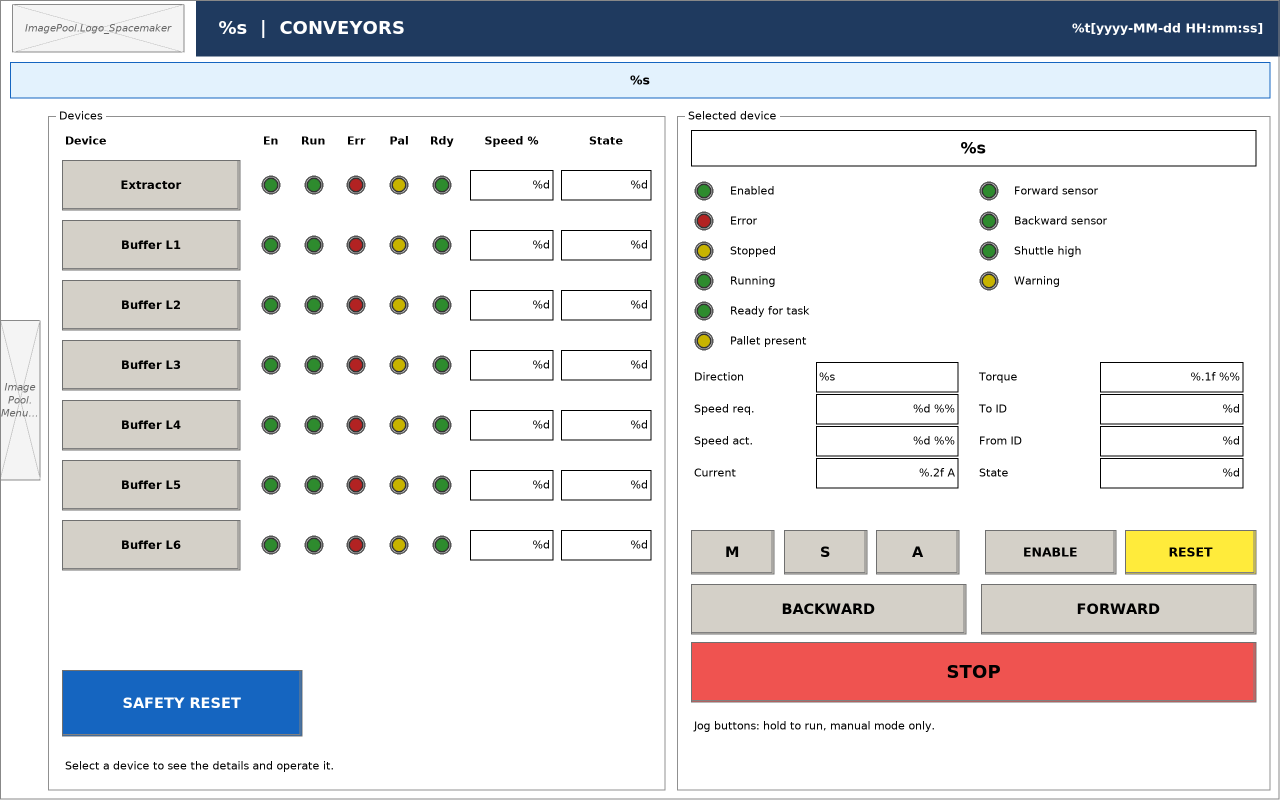
VISUALIZATION CNV  // 1280x800
    Rectangle (0,0 196x56)
        OnMouseClick: change screen: Main
    Image (12,4 172x48), image: ImagePool.Logo_Spacemaker
        OnMouseClick: change screen: Main
    Rectangle (196,0 1084x56), "%s | CONVEYORS", text variable: GVL_HMI_System.stStatus.sSystemName
    Rectangle (930,8 336x40), "%t[yyyy-MM-dd HH:mm:ss]", text variable: GVL_HMI_System.stStatus.dtNow
    Rectangle (10,62 1260x36), "%s", text variable: GVL_HMI_System.stStatus.sMessage, colour toggle: GVL_HMI_System.stStatus.bMessageAlarm
    GroupBox (48,108 617x682), "Devices"
    Rectangle (62,128 178x26), "Device"
    Rectangle (250,128 42x26), "En"
    Rectangle (292,128 43x26), "Run"
    Rectangle (335,128 43x26), "Err"
    Rectangle (378,128 43x26), "Pal"
    Rectangle (421,128 42x26), "Rdy"
    Rectangle (470,128 83x26), "Speed %"
    Rectangle (561,128 90x26), "State"
    Button (62,160 178x50), "Extractor", colour toggle: GVL_HMI_CNV.astConveyor[0].bSelected
        OnMouseClick: execute { GVL_HMI_CNV.uiSelected := 0; }
    Lamp1 (260,174 22x22), variable: GVL_HMI_CNV.astConveyor[0].bEnabled, style: Lamp-Lamp1-Green
    Lamp1 (303,174 22x22), variable: GVL_HMI_CNV.astConveyor[0].bRunning, style: Lamp-Lamp1-Green
    Lamp1 (345,174 22x22), variable: GVL_HMI_CNV.astConveyor[0].bError, style: Lamp-Lamp1-Red
    Lamp1 (388,174 22x22), variable: GVL_HMI_CNV.astConveyor[0].bOccupied, style: Lamp-Lamp1-Yellow
    Lamp1 (431,174 22x22), variable: GVL_HMI_CNV.astConveyor[0].bReadyForTask, style: Lamp-Lamp1-Green
    Rectangle (470,170 83x30), "%d", text variable: GVL_HMI_CNV.astConveyor[0].iSpeedActual_pct
    Rectangle (561,170 90x30), "%d", text variable: GVL_HMI_CNV.astConveyor[0].uiStateMachine
    Button (62,220 178x50), "Buffer L1", colour toggle: GVL_HMI_CNV.astConveyor[1].bSelected
        OnMouseClick: execute { GVL_HMI_CNV.uiSelected := 1; }
    Lamp1 (260,234 22x22), variable: GVL_HMI_CNV.astConveyor[1].bEnabled, style: Lamp-Lamp1-Green
    Lamp1 (303,234 22x22), variable: GVL_HMI_CNV.astConveyor[1].bRunning, style: Lamp-Lamp1-Green
    Lamp1 (345,234 22x22), variable: GVL_HMI_CNV.astConveyor[1].bError, style: Lamp-Lamp1-Red
    Lamp1 (388,234 22x22), variable: GVL_HMI_CNV.astConveyor[1].bOccupied, style: Lamp-Lamp1-Yellow
    Lamp1 (431,234 22x22), variable: GVL_HMI_CNV.astConveyor[1].bReadyForTask, style: Lamp-Lamp1-Green
    Rectangle (470,230 83x30), "%d", text variable: GVL_HMI_CNV.astConveyor[1].iSpeedActual_pct
    Rectangle (561,230 90x30), "%d", text variable: GVL_HMI_CNV.astConveyor[1].uiStateMachine
    Button (62,280 178x50), "Buffer L2", colour toggle: GVL_HMI_CNV.astConveyor[2].bSelected
        OnMouseClick: execute { GVL_HMI_CNV.uiSelected := 2; }
    Lamp1 (260,294 22x22), variable: GVL_HMI_CNV.astConveyor[2].bEnabled, style: Lamp-Lamp1-Green
    Lamp1 (303,294 22x22), variable: GVL_HMI_CNV.astConveyor[2].bRunning, style: Lamp-Lamp1-Green
    Lamp1 (345,294 22x22), variable: GVL_HMI_CNV.astConveyor[2].bError, style: Lamp-Lamp1-Red
    Lamp1 (388,294 22x22), variable: GVL_HMI_CNV.astConveyor[2].bOccupied, style: Lamp-Lamp1-Yellow
    Lamp1 (431,294 22x22), variable: GVL_HMI_CNV.astConveyor[2].bReadyForTask, style: Lamp-Lamp1-Green
    Rectangle (470,290 83x30), "%d", text variable: GVL_HMI_CNV.astConveyor[2].iSpeedActual_pct
    Rectangle (561,290 90x30), "%d", text variable: GVL_HMI_CNV.astConveyor[2].uiStateMachine
    Button (62,340 178x50), "Buffer L3", colour toggle: GVL_HMI_CNV.astConveyor[3].bSelected
        OnMouseClick: execute { GVL_HMI_CNV.uiSelected := 3; }
    Lamp1 (260,354 22x22), variable: GVL_HMI_CNV.astConveyor[3].bEnabled, style: Lamp-Lamp1-Green
    Lamp1 (303,354 22x22), variable: GVL_HMI_CNV.astConveyor[3].bRunning, style: Lamp-Lamp1-Green
    Lamp1 (345,354 22x22), variable: GVL_HMI_CNV.astConveyor[3].bError, style: Lamp-Lamp1-Red
    Lamp1 (388,354 22x22), variable: GVL_HMI_CNV.astConveyor[3].bOccupied, style: Lamp-Lamp1-Yellow
    Lamp1 (431,354 22x22), variable: GVL_HMI_CNV.astConveyor[3].bReadyForTask, style: Lamp-Lamp1-Green
    Rectangle (470,350 83x30), "%d", text variable: GVL_HMI_CNV.astConveyor[3].iSpeedActual_pct
    Rectangle (561,350 90x30), "%d", text variable: GVL_HMI_CNV.astConveyor[3].uiStateMachine
    Button (62,400 178x50), "Buffer L4", colour toggle: GVL_HMI_CNV.astConveyor[4].bSelected
        OnMouseClick: execute { GVL_HMI_CNV.uiSelected := 4; }
    Lamp1 (260,414 22x22), variable: GVL_HMI_CNV.astConveyor[4].bEnabled, style: Lamp-Lamp1-Green
    Lamp1 (303,414 22x22), variable: GVL_HMI_CNV.astConveyor[4].bRunning, style: Lamp-Lamp1-Green
    Lamp1 (345,414 22x22), variable: GVL_HMI_CNV.astConveyor[4].bError, style: Lamp-Lamp1-Red
    Lamp1 (388,414 22x22), variable: GVL_HMI_CNV.astConveyor[4].bOccupied, style: Lamp-Lamp1-Yellow
    Lamp1 (431,414 22x22), variable: GVL_HMI_CNV.astConveyor[4].bReadyForTask, style: Lamp-Lamp1-Green
    Rectangle (470,410 83x30), "%d", text variable: GVL_HMI_CNV.astConveyor[4].iSpeedActual_pct
    Rectangle (561,410 90x30), "%d", text variable: GVL_HMI_CNV.astConveyor[4].uiStateMachine
    Button (62,460 178x50), "Buffer L5", colour toggle: GVL_HMI_CNV.astConveyor[5].bSelected
        OnMouseClick: execute { GVL_HMI_CNV.uiSelected := 5; }
    Lamp1 (260,474 22x22), variable: GVL_HMI_CNV.astConveyor[5].bEnabled, style: Lamp-Lamp1-Green
    Lamp1 (303,474 22x22), variable: GVL_HMI_CNV.astConveyor[5].bRunning, style: Lamp-Lamp1-Green
    Lamp1 (345,474 22x22), variable: GVL_HMI_CNV.astConveyor[5].bError, style: Lamp-Lamp1-Red
    Lamp1 (388,474 22x22), variable: GVL_HMI_CNV.astConveyor[5].bOccupied, style: Lamp-Lamp1-Yellow
    Lamp1 (431,474 22x22), variable: GVL_HMI_CNV.astConveyor[5].bReadyForTask, style: Lamp-Lamp1-Green
    Rectangle (470,470 83x30), "%d", text variable: GVL_HMI_CNV.astConveyor[5].iSpeedActual_pct
    Rectangle (561,470 90x30), "%d", text variable: GVL_HMI_CNV.astConveyor[5].uiStateMachine
    Button (62,520 178x50), "Buffer L6", colour toggle: GVL_HMI_CNV.astConveyor[6].bSelected
        OnMouseClick: execute { GVL_HMI_CNV.uiSelected := 6; }
    Lamp1 (260,534 22x22), variable: GVL_HMI_CNV.astConveyor[6].bEnabled, style: Lamp-Lamp1-Green
    Lamp1 (303,534 22x22), variable: GVL_HMI_CNV.astConveyor[6].bRunning, style: Lamp-Lamp1-Green
    Lamp1 (345,534 22x22), variable: GVL_HMI_CNV.astConveyor[6].bError, style: Lamp-Lamp1-Red
    Lamp1 (388,534 22x22), variable: GVL_HMI_CNV.astConveyor[6].bOccupied, style: Lamp-Lamp1-Yellow
    Lamp1 (431,534 22x22), variable: GVL_HMI_CNV.astConveyor[6].bReadyForTask, style: Lamp-Lamp1-Green
    Rectangle (470,530 83x30), "%d", text variable: GVL_HMI_CNV.astConveyor[6].iSpeedActual_pct
    Rectangle (561,530 90x30), "%d", text variable: GVL_HMI_CNV.astConveyor[6].uiStateMachine
    Rectangle (62,752 593x28), "Select a device to see the details and operate it."
    GroupBox (677,108 593x682), "Selected device"
    Rectangle (691,130 565x36), "%s", text variable: GVL_HMI_CNV.stSelected.sName
    Lamp1 (693,180 22x22), variable: GVL_HMI_CNV.stSelected.bEnabled, style: Lamp-Lamp1-Green
    Rectangle (727,176 201x30), "Enabled"
    Lamp1 (693,210 22x22), variable: GVL_HMI_CNV.stSelected.bError, style: Lamp-Lamp1-Red
    Rectangle (727,206 201x30), "Error"
    Lamp1 (693,240 22x22), variable: GVL_HMI_CNV.stSelected.bStopped, style: Lamp-Lamp1-Yellow
    Rectangle (727,236 201x30), "Stopped"
    Lamp1 (693,270 22x22), variable: GVL_HMI_CNV.stSelected.bRunning, style: Lamp-Lamp1-Green
    Rectangle (727,266 201x30), "Running"
    Lamp1 (693,300 22x22), variable: GVL_HMI_CNV.stSelected.bReadyForTask, style: Lamp-Lamp1-Green
    Rectangle (727,296 201x30), "Ready for task"
    Lamp1 (693,330 22x22), variable: GVL_HMI_CNV.stSelected.bOccupied, style: Lamp-Lamp1-Yellow
    Rectangle (727,326 201x30), "Pallet present"
    Lamp1 (978,180 22x22), variable: GVL_HMI_CNV.stSelected.bForwardSensor, style: Lamp-Lamp1-Green
    Rectangle (1011,176 202x30), "Forward sensor"
    Lamp1 (978,210 22x22), variable: GVL_HMI_CNV.stSelected.bBackwardSensor, style: Lamp-Lamp1-Green
    Rectangle (1011,206 202x30), "Backward sensor"
    Lamp1 (978,240 22x22), variable: GVL_HMI_CNV.stSelected.bShuttleHigh, style: Lamp-Lamp1-Green
    Rectangle (1011,236 202x30), "Shuttle high"
    Lamp1 (978,270 22x22), variable: GVL_HMI_CNV.stSelected.bWarning, style: Lamp-Lamp1-Yellow
    Rectangle (1011,266 202x30), "Warning"
    Rectangle (691,362 119x30), "Direction"
    Rectangle (816,362 142x30), "%s", text variable: GVL_HMI_CNV.stSelected.sMotorDirection
    Rectangle (691,394 119x30), "Speed req."
    Rectangle (816,394 142x30), "%d %%", text variable: GVL_HMI_CNV.stSelected.iSpeedRequested_pct
    Rectangle (691,426 119x30), "Speed act."
    Rectangle (816,426 142x30), "%d %%", text variable: GVL_HMI_CNV.stSelected.iSpeedActual_pct
    Rectangle (691,458 119x30), "Current"
    Rectangle (816,458 142x30), "%.2f A", text variable: GVL_HMI_CNV.stSelected.rCurrent_A
    Rectangle (976,362 118x30), "Torque"
    Rectangle (1100,362 143x30), "%.1f %%", text variable: GVL_HMI_CNV.stSelected.rTorque_pct
    Rectangle (976,394 118x30), "To ID"
    Rectangle (1100,394 143x30), "%d", text variable: GVL_HMI_CNV.stSelected.diTransferToId
    Rectangle (976,426 118x30), "From ID"
    Rectangle (1100,426 143x30), "%d", text variable: GVL_HMI_CNV.stSelected.diTransferFromId
    Rectangle (976,458 118x30), "State"
    Rectangle (1100,458 143x30), "%d", text variable: GVL_HMI_CNV.stSelected.uiStateMachine
    Button (691,530 83x44), "M", colour toggle: GVL_HMI_CNV.stSelected.bModeManual
        tap GVL_HMI_CNV.stCommand.bModeManual p3779583253=TRUE
    Button (784,530 83x44), "S", colour toggle: GVL_HMI_CNV.stSelected.bModeSemi
        tap GVL_HMI_CNV.stCommand.bModeSemi p3779583253=TRUE
    Button (876,530 83x44), "A", colour toggle: GVL_HMI_CNV.stSelected.bModeAuto
        tap GVL_HMI_CNV.stCommand.bModeAuto p3779583253=TRUE
    Button (985,530 131x44), "ENABLE", colour toggle: GVL_HMI_CNV.stSelected.bEnabled
        tap GVL_HMI_CNV.stCommand.bEnable p3779583253=TRUE
    Button (1125,530 131x44), "RESET"
        tap GVL_HMI_CNV.stCommand.bReset p3779583253=TRUE
    Button (691,584 275x50), "BACKWARD", input disabled if: NOT GVL_HMI_CNV.stSelected.bModeManual
        tap GVL_HMI_CNV.stCommand.bJogBackward p3779583253=TRUE
    Button (981,584 275x50), "FORWARD", input disabled if: NOT GVL_HMI_CNV.stSelected.bModeManual
        tap GVL_HMI_CNV.stCommand.bJogForward p3779583253=TRUE
    Button (691,642 565x60), "STOP"
        tap GVL_HMI_CNV.stCommand.bStop p3779583253=TRUE
    Rectangle (691,712 565x28), "Jog buttons: hold to run, manual mode only."
    Rectangle (0,320 40x160)
        OnMouseClick: OpenDialog Dialog=Dialog, OpenModal=True, PositionX=0, PositionY=0
        OnMouseEnter: OpenDialog Dialog=Dialog, OpenModal=True, PositionX=0, PositionY=0
    Image (0,320 40x160), image: ImagePool.Menu_Tab
        OnMouseClick: OpenDialog Dialog=Dialog, OpenModal=True, PositionX=0, PositionY=0
        OnMouseEnter: OpenDialog Dialog=Dialog, OpenModal=True, PositionX=0, PositionY=0
    Button (62,670 240x66), "SAFETY RESET", colour toggle: GVL_HMI_System.stStatus.bSafetyResetActive
        tap GVL_HMI_System.stCommand.bSafetyReset p3779583253=TRUE
END_VISUALIZATION

(* stored: Version 1.1.0.1
   Visu CNV: Id {bd5207fc-b697-4aa5-9856-89eae20f8f06} *)
